// TIA Portal V21 export
// export: Created 2026-11-10T07:27:00.4231252Z, ExportSetting WithDefaults, DisplayName Totally Integrated Automation Portal, DisplayVersion V21 Update 3, DisplayName STEP 7 Professional, DisplayVersion V21 Update 3, DisplayName STEP 7 Safety, DisplayVersion V21, DisplayName Tech WebApplication, DisplayVersion V21, DisplayName WinCC Basic/Comfort/Advanced, DisplayVersion V21 Update 3, DisplayName WinCC Unified, DisplayVersion V21 Update 3
FUNCTION "FC_SclRest" : Void   // FC14, SCL
{ S7_Optimized_Access := 'TRUE' }
VERSION : 0.1
// stored: AutoNumber true, IsIECCheckEnabled false, SetENOAutomatically false, UDAEnableTagReadback false
   VAR_INPUT
      anyp : Any;
      ptrp : Pointer;
      sp : Real;
   END_VAR
   VAR_TEMP
      x : Int;
      y : Int;
      "b" : Bool;
      "by" : Byte;
      w : Word;
      dw : DWord;
      rp : REF_TO Int;
      rd : REF_TO "UDT_Motor";
      v : Variant;
   END_VAR
BEGIN
   // peek and poke variants
   #by := PEEK(area := 16#84, dbNumber := 1, byteOffset := 0);
   #w := PEEK_WORD(area := 16#84, dbNumber := 1, byteOffset := 0);
   #dw := PEEK_DWORD(area := 16#84, dbNumber := 1, byteOffset := 0);
   #b := PEEK_BOOL(area := 16#84, dbNumber := 1, byteOffset := 0, bitOffset := 1);
   POKE(area := 16#84, dbNumber := 1, byteOffset := 0, value := #by);
   POKE(area := 16#84, dbNumber := 1, byteOffset := 0, value := #w);
   POKE(area := 16#84, dbNumber := 1, byteOffset := 0, value := #dw);
   POKE_BOOL(area := 16#84, dbNumber := 1, byteOffset := 0, bitOffset := 1, value := #b);
   // references and dereferencing
   #rp := REF("DB_Global".iInt);
   #rp^ := 5;
   #y := #rp^;
   #b := #rp = NULL;
   #b := #rp <> NULL;
   #rd := REF("DB_Motor".motor);
   #y := #rd^.Count;
   // absolute DB address with explicit bit
   "DB_Std".x := TRUE;
END_FUNCTION
